# EPICS autosave request: utcaApp/Db/pbpm_pos_calc.req
$(P)$(R)PosKx-SP
$(P)$(R)PosKy-SP
$(P)$(R)SupMat-SP
$(P)$(R)PosXOffset-SP
$(P)$(R)PosYOffset-SP
